TYPE ST_PERIPHERY_REF : FB_PERIPHERY_REF;
END_TYPE

(* stored: Version 1.1.0.1, ProductVersion 3.1.4024.15
   DUT ST_PERIPHERY_REF: Id {3d1c9026-b3b6-4865-ad38-a21940b7764a} *)
